(* IEC 61131-3 sources: PortalRobot/Portal_robot/Device/application/ST/ST_ALARM, 10 files *)

(* ---- E_ALARM_EFFECT.st ---- *)
TYPE E_ALARM_EFFECT :
(
	GLOBAL_STOP, // Аварийный останов всей ячейки
	ROBOT_STOP, // Останов робота и текущего взаимодействия с оборудованием
	EQUIPMENT_STOP, // Останов только владельца аварии
	WARNING // Информационное предупреждение без останова
);
END_TYPE

(* ---- E_ALARM_SEVERITY.st ---- *)
TYPE E_ALARM_SEVERITY :
(
	ALARM, // Авария, требующая устранения причины
	WARNING // Предупреждение оператору
);
END_TYPE

(* ---- E_ALARM_SOURCE.st ---- *)
TYPE E_ALARM_SOURCE :
(
	CELL, // Ячейка
	ROBOT, // Робот
	MACHINE_1, // Станок 1
	MACHINE_2, // Станок 2
	MACHINE_3, // Станок 3
	MAGAZINE_LOGIC_1, // Магазин 1; имя не конфликтует с SoftMotion-осью Magazine_1
	MAGAZINE_LOGIC_2, // Магазин 2; имя не конфликтует с SoftMotion-осью Magazine_2
	RESERVED_LEGACY_MAGAZINE_AXIS_1, // Код 7 сохранён только для старых записей журнала
	RESERVED_LEGACY_MAGAZINE_AXIS_2, // Код 8 сохранён только для старых записей журнала
	AXIS_X, // Ось X
	AXIS_Y, // Ось Y
	AXIS_Z, // Ось Z
	AXIS_GROUP, // Группа осей XYZ
	MOTION_MANAGER, // Менеджер движения
	POINT_MANAGER, // Менеджер точек
	GRIPPER, // Захват робота
	CELL_SAFETY, // Дискретный контур безопасности; прежние числовые коды сохранены
	GEOMETRY_1,
	GEOMETRY_2,
    CONTROLLER_CPU_1, // Коды 19..21 добавлены без изменения прежней нумерации.
    CONTROLLER_CPU_2,
    CONTROLLER_MODULES
);
END_TYPE

(* ---- ST_ALARM_COMMAND.st ---- *)
TYPE ST_ALARM_COMMAND :
STRUCT
	xResetWarnings : BOOL; // Импульс сброса накопленных предупреждений
END_STRUCT
END_TYPE

(* ---- ST_ALARM_EVENT.st ---- *)
TYPE ST_ALARM_EVENT :
STRUCT
	udiSequence : UDINT; // Уникальный порядковый номер события
	eSeverity   : E_ALARM_SEVERITY; // Уровень события
	eEffect     : E_ALARM_EFFECT; // Фактическое воздействие события в момент фиксации
	eSource     : E_ALARM_SOURCE; // Механизм-источник события
	uiCode      : UINT; // Номер бита ошибки или код предупреждения
	xActive     : BOOL; // Событие ещё активно и требует внимания
END_STRUCT
END_TYPE

(* ---- ST_ALARM_SOURCE_DATA.st ---- *)
TYPE ST_ALARM_SOURCE_DATA :
STRUCT
	eSource       : E_ALARM_SOURCE; // Функциональный блок, которому принадлежит событие
	dwAlarmActive : DWORD; // Только собственные активные аварии блока
	xRobotStopRequired : BOOL; // Владелец зафиксировал зависимый останов робота для этого контекста
	xGlobalError  : BOOL; // Глобальная ошибка была активна в момент публикации источника
	stWarning     : ST_WARNING_EVENT; // Последнее предупреждение блока
END_STRUCT
END_TYPE

(* ---- ST_ALARM_STATUS.st ---- *)
TYPE ST_ALARM_STATUS :
STRUCT
	uiActiveAlarmCount   : UINT; // Число активных аварий
	uiActiveWarningCount : UINT; // Число активных предупреждений
	uiActiveEventCount   : UINT; // Общее число активных событий
	uiHistoryCount       : UINT; // Число записей в журнале
	xAlarmActive         : BOOL; // Есть хотя бы одна активная авария
	xWarningActive       : BOOL; // Есть хотя бы одно активное предупреждение
END_STRUCT
END_TYPE

(* ---- ST_CONTROLLER_WEB_REQUEST.st ---- *)
TYPE ST_CONTROLLER_WEB_REQUEST :
STRUCT
    udiSequence : UDINT; // Gateway записывает последним; payload неизменен до Ack.
    udiIssuedAtMs : UDINT; // Часы PLC, прочитанные перед передачей.
    xCpuValid : BOOL;
    xModulesValid : BOOL;
    dwCpuCurrent1 : DWORD;
    dwCpuCurrent2 : DWORD;
    dwModuleCurrent : DWORD;
    xMemoryCurrent : BOOL;
    dwCpuObserved1 : DWORD; // Причины, обнаруженные с прошлого подтверждения PLC.
    dwCpuObserved2 : DWORD;
    dwModuleObserved : DWORD;
    xMemoryObserved : BOOL;
END_STRUCT
END_TYPE

(* ---- ST_CONTROLLER_WEB_STATUS.st ---- *)
TYPE ST_CONTROLLER_WEB_STATUS :
STRUCT
    udiAckSeq : UDINT;
    dwCpuAlarm1 : DWORD;
    dwCpuAlarm2 : DWORD;
    dwModuleAlarm : DWORD;
    xMemoryWarning : BOOL;
    xCpuFresh : BOOL;
    xModulesFresh : BOOL;
    xAlarmActive : BOOL;
    xGlobalStopRequired : BOOL;
    xResetAllowed : BOOL;
    xWarningResetAllowed : BOOL;
END_STRUCT
END_TYPE

(* ---- ST_WARNING_EVENT.st ---- *)
TYPE ST_WARNING_EVENT :
STRUCT
	udiSequence : UDINT; // Порядковый номер предупреждения от функционального блока
	uiCode      : UINT; // Код предупреждения внутри функционального блока
END_STRUCT
END_TYPE
